      if get_inverse_kin_has_solution(pose.crt, qnear=pose.q):
          pose.jnt = get_inverse_kin(pose.crt, qnear=pose.q)
      else:
          popup("no solution found for the transition pose", blocking= True)
      end

      return pose
  end

  def get_transition_pose_2(ref, radius, axis_config, closest=False):
      # get the correspondig pose from the list of poses

      local jnt_current = get_actual_joint_positions()
      local yaw_current = get_yaw_too_base(ref)

      #pose.crt = get_tool_free_pose(pose_ref=ref, dir=[0, 0, DISTANCE_TO_CLEARANCE], move_in_base_frame=True)

      if (axis_config == 1):
          pose.q = JNT_STANDARD_C1
      elif (axis_config == 2):
          pose.q = JNT_STANDARD_C2
      end

      if closest:
          pose.q[0] = jnt_current[0]
      end

      # get coordinates of the circle with the same angle as the given pose to the
      if ref == p[0,0,0,0,0,0]:
          pose.crt = PSE_WA_1
      else:
          pose.crt =
          p[radius * cos(yaw_current-pi/2),
          radius * sin(yaw_current-pi/2),
          DISTANCE_TO_CLEARANCE,
          0,
          0,
          yaw_current + get_locked_yaw()]
      end

      if get_inverse_kin_has_solution(pose.crt, qnear=pose.q):
          pose.jnt = get_inverse_kin(pose.crt, qnear=pose.q)
          #return pose
      else:
          popup("no solution found for the transition pose", blocking= True)
      end

      return pose
  end

  def get_rounded_mm(value):
      if (value < 0):
          return ceil(value*1000)
      elif (value >= 0):
          return floor(value*1000)
      end
  end

  def get_yaw_too_base(pose):
      # get the yaw relative to the base frame
      local pose_x_mm = 0
      local pose_y_mm = 0
      local yaw = 0

      pose_x_mm = get_rounded_mm(pose[0])
      pose_y_mm = get_rounded_mm(pose[1])

      if (pose_x_mm == 0 and pose_y_mm < 0):
          yaw = 0
      elif (pose_x_mm == 0 and pose_y_mm > 0):
          yaw = pi
      elif (pose_x_mm < 0 and pose_y_mm == 0):
          yaw = -pi/2
      elif (pose_x_mm > 0 and pose_y_mm == 0):
          yaw = pi/2
      else:
          yaw = atan2(pose[0], pose[1])
          if (-pi < yaw) and (yaw < 0):
              yaw = - yaw - pi
          elif (0 < yaw) and (yaw < pi):
              yaw = - yaw + pi
          else:
              yaw = pi
          end
      end
      return yaw
  end

  def get_helper_pose():
      # get the helper pose, as described

      local m_line = 0                    # slope of the line between base and circle point
      local n = 0                         # shift on the ordinate axis
      local m_normal = 0                  # slope of the normal of the line between base and circle point
      local x_p1 = 0                      # x coordinate of first circle point
      local x_p2 = 0                      # x coordinate of second circle point
      local y_p1 = 0                      # y coordinate of first circle point
      local y_p2 = 0                      # y coordinate of second circle point
      local jnt_help_1 = [0,0,0,0,0,0]
      local jnt_help_2 = [0,0,0,0,0,0]

      if (pose_start.crt != pose_target.crt):
          if (pose_start.crt[0] == pose_target.crt[0]):
              m_normal = 0
          elif (pose_start.crt[0] != pose_target.crt[0]):
              m_line = (pose_target.crt[1]-pose_start.crt[1])/(pose_target.crt[0]-pose_start.crt[0])    # calculation of the slope between start and target
              n = pose_start.crt[1] - m_line * pose_start.crt[0]
          end
          if (-0.00001 > m_line or m_line > 0.00001):
              m_normal = -1/m_line
          end

          # using p-q-formula for getting the crossing points
          x_p1 = sqrt(pow(RADIUS_HELPER_POSES, 2)/(pow(m_normal, 2)+1)) * -1
          x_p2 = sqrt(pow(RADIUS_HELPER_POSES, 2)/(pow(m_normal, 2)+1))
          y_p1 = m_normal * x_p1
          y_p2 = m_normal * x_p2
          pose.q = pose_start.jnt

          if (point_dist(pose_start.crt, p[x_p1, y_p1,0,0,0,0]) < point_dist(pose_start.crt, p[x_p2, y_p2,0,0,0,0])):
              if reverse_rotation:
                  pose_help.crt[0] = x_p2
                  pose_help.crt[1] = y_p2
                  pose.q = pose_target.jnt
              else:
                  pose_help.crt[0] = x_p1
                  pose_help.crt[1] = y_p1
                  pose.q = pose_start.jnt
              end
          elif (point_dist(pose_start.crt, p[x_p1, y_p1,0,0,0,0]) > point_dist(pose_start.crt, p[x_p2, y_p2,0,0,0,0])):
              if reverse_rotation:
                  pose_help.crt[0] = x_p1
                  pose_help.crt[1] = y_p1
                  pose.q = pose_target.jnt
              else:
                  pose_help.crt[0] = x_p2
                  pose_help.crt[1] = y_p2
                  pose.q = pose_start.jnt
              end
          elif (point_dist(pose_start.crt, p[x_p1, y_p1,0,0,0,0]) == point_dist(pose_start.crt, p[x_p2, y_p2,0,0,0,0])):
              jnt_help_1 = get_inverse_kin(p[x_p1, y_p1,pose_start.crt[2],pose_start.crt[3],pose_start.crt[4],pose_start.crt[5]], qnear=pose.q)
              jnt_help_2 = get_inverse_kin(p[x_p2, y_p2,pose_start.crt[2],pose_start.crt[3],pose_start.crt[4],pose_start.crt[5]], qnear=pose.q)
              if (pose_start.jnt[0]<jnt_help_1[0] and jnt_help_1[0]<pose_target.jnt[0]) or (pose_start.jnt[0]>jnt_help_1[0] and jnt_help_1[0]>pose_target.jnt[0]):
                  pose_help.crt[0] = x_p1
                  pose_help.crt[1] = y_p1
              elif (pose_start.jnt[0]<jnt_help_2[0] and jnt_help_2[0]<pose_target.jnt[0]) or (pose_start.jnt[0]>jnt_help_2[0] and jnt_help_2[0]>pose_target.jnt[0]):
                  pose_help.crt[0] = x_p2
                  pose_help.crt[1] = y_p2
              end
              pose.q = pose_start.jnt
          end

          pose_help.crt[2] = 0.5 * (pose_start.crt[2] + pose_target.crt[2])

          if ((pose_start.crt[1] < 0 and pose_target.crt[1] > 0) or (pose_start.crt[1] > 0 and pose_target.crt[1] < 0)):
              if get_inverse_kin_has_solution(pose.crt, qnear=pose.q):
                  pose.jnt = get_inverse_kin(pose.crt, qnear=pose.q)
              else:
                  popup("no solution found for the helper pose", blocking= True)
              end
          end
      end
      return pose
  end

  def adjust_transition_poses(pose_identifier):
      # adjust the orientation of the transition poses by determining the the current orientation

      local pose_current = get_actual_tcp_pose()
      local jnt_current = get_actual_joint_positions()
      local rpy_current = rotvec2rpy([pose_current[3],pose_current[4],pose_current[5]])
      local rotvec_new = [0,0,0]

      if (pose_identifier == "start"):
          pose.q = pose_start.jnt
          pose.crt = get_forward_kin(pose_start.jnt)
      elif (pose_identifier == "helper"):
          pose.q = pose_help.jnt
          pose.crt = get_forward_kin(pose_help.jnt)
      elif (pose_identifier == "target"):
          pose.q = pose_target.jnt
          pose.crt = get_forward_kin(pose_target.jnt)
      end

      rotvec_new = rpy2rotvec([rpy_current[0], rpy_current[1], get_yaw_too_base(pose.crt) + yaw_locked])
      pose.crt = p[pose.crt[0], pose.crt[1], pose.crt[2], rotvec_new[0], rotvec_new[1], rotvec_new[2]]

      pose.q[3] = jnt_current[3]
      pose.q[4] = jnt_current[4]
      pose.q[5] = jnt_current[5]
      if get_inverse_kin_has_solution(pose.crt, qnear=pose.q) and is_within_safety_limits(pose.crt):
          pose.jnt = get_inverse_kin(pose.crt, qnear=pose.q)
      else:
          popup(str_cat("no solution for ", pose_identifier), error=True, blocking=True)
      end
      return pose.jnt
  end

  def get_locked_yaw():
      local pose_current = get_actual_tcp_pose()
      local rpy_current = rotvec2rpy([pose_current[3],pose_current[4],pose_current[5]])
      local rotvec_new = rpy2rotvec([rpy_current[0], rpy_current[1], get_yaw_too_base(pose_current)])
      local pose_reference = p[pose_current[0], pose_current[1], pose_current[2], rotvec_new[0], rotvec_new[1], rotvec_new[2]]
      local pose_to_reference = pose_trans(pose_inv(pose_reference), get_actual_tcp_pose())
      yaw_locked = pose_to_reference[5]

      return yaw_locked
  end

  def do_transition(reference_pose=p[0,0,0,0,0,0], mode=2, keep_xyz=[False, False, False], keep_rxry=False, a=1.4, v=1.05, r=0.100):
      # the robot will evaluate the current and target workarea
      # after that, the robot will move between the workareas automatically.
      # parameters:
      # reference_pose:   a pose/frame were the robot should work next. If nothing is given, base frame will be used as target
      # keep_rxry:        if true, the robot will keep the orientation of the tool during the movement

      ################# checking #################
      axis_config_current = check_current_axis_config()           # 0: unknown, 1: config 1, 2: config 2
      workarea_current = check_workarea(get_actual_tcp_pose())    # between 0 and the amount of defined workareas
      workarea_new = check_workarea(reference_pose)               # between 0 and the amount of defined workareas
      if(workarea_current==workarea_new):
           return 0
      end
      if (workarea_current != 0 and workarea_new != 0):
          ################# get axisvalues #################
          # pose_start = get_transition_pose(workarea_current, axis_config_current, closest=not reverse_rotation, keep_xyz=keep_xyz)
          pose_start = get_transition_pose_2(get_actual_tcp_pose(), RADIUS_TRANSITION_POSES, axis_config_current, closest=not reverse_rotation)
          if (workarea_current == 3 and workarea_new == 4) or (workarea_current == 4 and workarea_new == 3):
              # pose_target = get_transition_pose(workarea_new, axis_config_current, closest=True)
              pose_target = get_transition_pose_2(reference_pose, RADIUS_TRANSITION_POSES, axis_config_current, closest=True)
              reverse_rotation = True
          else:
              pose_target = get_transition_pose_2(reference_pose, RADIUS_TRANSITION_POSES, axis_config_current, closest=(workarea_current == workarea_new))
              if reverse_rotation:
                  reverse_rotation = False
              end
          end
          # pose_help = get_helper_pose()
          global A_Start = pose_start.crt
          global A_Help = pose_help.crt
          global A_End = pose_target.crt


          ################# adjustments #################
          if (keep_rxry):
              get_locked_yaw()
              if (pose_start.jnt == pose_target.jnt):
                  pose_target.jnt = adjust_transition_poses("target")
                  pose_start.jnt = pose_target.jnt
              else:
                  pose_start.jnt = adjust_transition_poses("start")
                  pose_target.jnt = adjust_transition_poses("target")
              end
              if (pose_help.jnt != [0,0,0,0,0,0]):
                  pose_help.jnt = adjust_transition_poses("helper")
              end
          end

          global A_Start = pose_start.crt
          global A_Help = pose_help.crt
          global A_End = pose_target.crt

          ################# movements #################

          if point_dist(pose_start.crt, pose_target.crt) > 0.100:
              movej(pose_start.jnt, a=a, v=v, r=r)
          end
          # if (pose_help.jnt != [0,0,0,0,0,0]):
          #     movej(pose_help.jnt, a=a, v=v, r=r)
          # end
          movej(pose_target.jnt, a=a, v=v)
      else:
          # define error
      end

      ################# checking #################
      axis_config_current = check_current_axis_config()           # 0: unknown, 1: config 1, 2: config 2
      workarea_current = check_workarea(get_actual_tcp_pose())    # between 0 and the amount of defined workareas
  end
  $ 5 "Script: SCRIPT Utility V5.1.script"
  #*****************************************************
  # customer          :   tbd
  # project name      :   tbd
  #****************************************************
  # controller        :
  # software          :
  #****************************************************
  # author            :   P. Koehnke (+49 1628859904; p.koehnke@unitedrobotics.group)
  # Copyright (c)     :   United Robotics Group Health and Food GmbH
  #                       An der Riede 2
  #                       28816 Stuhr
  #                       Germany
  #****************************************************
  # description       :   utility programs for the application
  # version:      	:   3.1
  # created           :   30.01.2023
  # updated           :
  #****************************************************
  # modifications     :   get_tool_free_pose_2(), get_index_from_list()
  #
  # date              :   05.01.2024
  # name              :   PK
  # reason            :
  #****************************************************

  def found_in_matrix(data, req_id, req_idx):
      local id = -1
      local dimensions = size(data)
      local loop_dataset = 0

      while (id != req_id and loop_dataset < dimensions[0]):
          id = data[loop_dataset, 0]
          if (id == req_id):
              return data[loop_dataset, req_idx]
          else:
              loop_dataset = loop_dataset + 1
          end
      end
  end

  def found_in_list(value, list):
      local idx = 0

      while (idx < length(list)):
          if (value == list[idx]):
              return True
          end
          idx = idx + 1
      end
      return False
  end

  def get_index_from_list(list, value=-1):
      local idx = 0

      while (idx < length(list)):
          if (value == -1):
              if (list[idx] != 0):
                  return idx
              end
          else:
              if (list[idx] == value):
                  return idx
              end
          end
          idx = idx + 1
      end
      return -1
  end

  def pose_RPY2RotVec(pose):
      local rotvec = rpy2rotvec([d2r(pose[3]),d2r(pose[4]),d2r(pose[5])])
      return p[pose[0],pose[1],pose[2],rotvec[0],rotvec[1],rotvec[2]]
  end

  def pose_RotVec2RPY(pose):
      local rpy = rotvec2rpy([pose[3],pose[4],pose[5]])
      return p[pose[0],pose[1],pose[2],r2d(rpy[0]),r2d(rpy[1]),r2d(rpy[2])]
  end

  def swivel(frame_ref, angles=[0,0,0], pose=p[0,0,0,0,0,0]):

      local rpy_ref = [0,0,0]
      local rpy_new = [0,0,0]
      local rotvec_new = [0,0,0]
      local pose_from = p[0,0,0,0,0,0]
      local pose_to = p[0,0,0,0,0,0]
      local i = 0

      if (pose == p[0,0,0,0,0,0]):
          pose_to = pose_trans(pose_inv(frame_ref), get_actual_tcp_pose())
      else:
          pose_to = pose
      end

      rpy_ref = rotvec2rpy(frame_ref[3], frame_ref[4], frame_ref[5])

      while (i < 3):
          rpy_new[i] = rpy_ref[i] + d2r(angles[i])
          i = i + 1
      end

      rotvec_new = rpy2rotvec(rpy_new)
      pose_from = p[0,0,0,rotvec_new[0],rotvec_new[1],rotvec_new[2]]
      pose_to = p[pose_to[0], pose_to[1], pose_to[2], rotvec_new[0], rotvec_new[1], rotvec_new[2]]

      return pose_trans(pose_from, pose_to)
  end

  def get_random_pose(pose_ref, mode="", range_max=[0,0,0]):
      # modi: "cubic", "rotation"
      # getting a random pose in the x/y-plane. range can be set for each
      # translation and rotation.
      local rpy_random = [0,0,0]
      local rotvec_random = [0,0,0]
      local pose_random = pose_ref
      local i = 0

      if (mode == "cubic"):
          # cubic mode: random pose takes only x, y and z
          i = 0
          while(i<3):
              pose_random[i] = pose_ref[i] + range_max[i] * (random() - 0.5)
              i = i + 1
          end
          return pose_random

      elif (mode == "rotation"):
          i = 0
          while(i<3):
              rpy_random[i] = d2r(range_max[i]) * (random() - 0.5)
              i = i + 1
          end
          rotvec_random = rpy2rotvec(rpy_random)
          pose_random = pose_trans(p[0,0,0,rotvec_random[0],rotvec_random[1],rotvec_random[2]], pose_ref)
          return pose_random

      else:
          # unknown mode, return pose_ref
          return pose_ref
      end
  end

  def get_pattern_pos_rectangle(counter, direction, patternsize, patterninc=[0,0], patternwidth=[0,0]):
      # defines the position inside a rectangular pattern
      # patternsize describes, how many objects are in x-direction and how many in y-direction [x, y]
      # patternwidth will give the total length of each direction [x, y]
      local X_Fac = 0
      local Y_Fac = 0
      local max = patternsize[0]*patternsize[1]

      if (1>counter or counter>max):
          counter = 1
      end

      if (direction == "Y" or direction == "y"):
          X_Fac = floor((counter - 1) / patternsize[1])
          Y_Fac = (counter - 1) % patternsize[1]
      elif (direction == "X" or direction == "x"):
          X_Fac = (counter - 1) % patternsize[0]
          Y_Fac = floor((counter - 1) / patternsize[0])
      end

      if patternwidth != [0,0]:
          patterninc = [patternwidth[0]/(patternsize[0]-1), patternwidth[1]/(patternsize[1]-1)]
      end

      return p[X_Fac*patterninc[0], Y_Fac*patterninc[1],0,0,0,0]
  end

  def get_pattern_pos_circle(counter, radius, angle, direction, pattern, patternsize=[0,0]):
      # get the patternpos for a circular pattern through a counter
      # need the radius and the angle in radiants
      local X_Fac = 0
      local Y_Fac = 0
      local rad_bow = 0
      local radius_cal = 0
      local ref = p[0,0,0,0,0,0]

      if (direction == "Y" or direction == "y"):
          X_Fac = floor((counter - 1) / pattern[1])
          Y_Fac = (counter - 1) % pattern[1]
      elif (direction == "X" or direction == "x"):
          X_Fac = (counter - 1) % pattern[0]
          Y_Fac = floor((counter - 1) / pattern[0])
      end

      # the opening angle will be calculated in x-direction
      # works only between -90 and 90 degree
      rad_bow = -angle/(pattern[0]-1) * X_Fac + angle/2

      if (counter%2 == 0):
          radius_cal = radius - patternsize[1]/(pattern[1])
      else:
          radius_cal = radius + patternsize[1]/(pattern[1])
      end
      ref = p[0, radius_cal, 0, 0, 0, 0]

      return p[ref[0]*cos(rad_bow)-ref[1]*sin(rad_bow), (ref[0]*sin(rad_bow)+ref[1]*cos(rad_bow))-radius,0,0,0,0]
  end

  def get_pattern_counter(pose, direction, pattern, patterninc=[0,0], patternsize=[0,0]):
      # returns the counter for a pattern from a given cartesian pose
      local patternpose = p[pose[0],pose[1],0,0,0,0]
      local floatFacX = 0.0
      local floatFacY = 0.0
      local remainder = 0.0
      local FacX = 0
      local FacY = 0

      # since the pattern spreads from the origin in positive axis-directions, all negative values
      # (which could appear due to a position near an axis) will set to zero
      if (pose[0]<0):
          patternpose = p[0,pose[1],0,0,0,0]
      end
      if (pose[1]<0):
          patternpose = p[pose[0],0,0,0,0,0]
      end
      # calculate the factor for each axis
      floatFacX = patternpose[0]/(patternsize[0]*(pattern[0]-1))
      floatFacY = patternpose[1]/(patternsize[1]*(pattern[1]-1))
      # determine the remainder after the comma/point
      if (floatFacX>1):
          remainder = floatFacX%floor(floatFacX)
      else:
          remainder = floatFacX
      end
      if (remainder<0.5):
          FacX = floatFacX-remainder
      else:
          FacX = floatFacX+(1-remainder)
      end

      if (floatFacY>1):
          remainder = floatFacY%floor(floatFacY)
      else:
          remainder = floatFacY
      end
      if (remainder<0.5):
          FacY = floatFacY-remainder
      else:
          FacY = floatFacY+(1-remainder)
      end
      # calculation of the counter in the desired axis-direction
      if (direction=="x" or direction=="X"):
          return FacX*pattern[1] + FacY + 1
      elif (direction=="y" or direction=="Y"):
          return FacY*pattern[0] + FacX + 1
      end
  end

  def get_plc_reg(mod_sig_name):
  	return integer_to_binary_list(modbus_get_signal_status(mod_sig_name))
  end

  def set_plc_reg(mod_sig_name, mod_sig_list):
  	modbus_set_output_register(mod_sig_name,binary_list_to_integer(mod_sig_list),False)
  end

  def check_decapping(offset=0, timeout=5):
      # checken, ob der Deckel schon ab ist
      local start = get_actual_tcp_pose()
      local current_offset = 0
      local timecounter = 0
      while (current_offset < offset):
          current_offset = pose_dist(start, get_actual_tcp_pose())
          timecounter = timecounter + 1
          if (timecounter*0.5 == timeout):
              break
          end
          sleep(0.5)
      end
      stopl(0.5)
  end

  def check_capping(torque=0):
      # checken, wann der Deckel verschraubt ist
      force_mode(get_actual_tcp_pose(), [0,0,1,0,0,0], [0,0,-2.0,0,0,0], 2, [0,0,0.100,0,0,0])
  end

  def is_reachable(frame, poses, offsets=[0,0,0]):
      local idx = 0
      local pose = p[0,0,0,0,0,0]

      while (idx < length(poses)):
          pose = poses[idx]
          pose[0] = pose[0] + offsets[0]
          pose[1] = pose[1] + offsets[1]
          pose[2] = pose[2] + offsets[2]

          if pose != p[0,0,0,0,0,0]:
              if (not get_inverse_kin_has_solution(pose_trans(frame, pose))):
                  textmsg(str_cat(str_cat("Pose ", to_str(idx + 1)), " is not reachable"))
                  return False
              end
          end
          idx = idx + 1
      end
      return True
  end

  def is_within_limits(frame, poses, offsets=[0,0,0]):
      local idx = 0
      local pose = p[0,0,0,0,0,0]

      while (idx < length(poses)):
          pose = poses[idx]
          pose[0] = pose[0] + offsets[0]
          pose[1] = pose[1] + offsets[1]
          pose[2] = pose[2] + offsets[2]

          if is_reachable(frame=frame, poses=poses, offsets=offsets):
              if (not is_within_safety_limits(get_inverse_kin(pose_trans(frame, pose), get_actual_joint_positions()))):
                  textmsg(str_cat(str_cat("Pose ", to_str(idx + 1)), "is out of joint limits"))
                  return False
              else:
                  idx = idx + 1
              end
          else:
              return False
          end
      end
      return True
  end

  def action_manipulator_decapping():
    zero_ftsensor()
    local DCP_Start = get_actual_tcp_pose ()
    global DCP_Actual = get_actual_tcp_pose ()
    local DCP_Height = 0.021
    global ForceCounter = 0
    sleep(0.02)
    zero_ftsensor()
    force_mode(p[0.0, 0.0, 0.0, 0.0, 0.0, 0.0], [0, 0, 1, 0, 0, 0], [0.0, 0.0, 17.0, 0.0, 0.0, 10.0], 2, [0.1, 0.1, 0.02, 0.3490658503988659, 0.3490658503988659, 0.3490658503988659])
    thread Thread_while_684():
      while (True):
        global DCP_Actual = get_actual_tcp_pose ()
        sleep(0.2)
        global ForceCounter = ForceCounter + 1
        if (ForceCounter > 30):
          zero_ftsensor()
          global ForceCounter = 0
        end
      end
    end
    if (DCP_Actual[2] <= DCP_Start[2] + DCP_Height):
      global thread_handler_decapping = run Thread_while_684()
      while (DCP_Actual[2] <= DCP_Start[2] + DCP_Height):
        sync()
      end
      kill thread_handler_decapping
    end
    end_force_mode()
    stopl(5.0)
  end
  $ 6 "PRC_Target≔0"
  global PRC_Target=0
  $ 7 "PRC_Target≔1"
  global PRC_Target=1
  $ 8 "Action≔1"
  global Action=1
  $ 9 "Action≔2"
  global Action=2
  $ 10 "Action≔7"
  global Action=7
  $ 11 "ITM_ID≔2"
  global ITM_ID=2
  $ 12 "JIG≔1"
  global JIG=1
  $ 13 "JIG_Slot≔2"
  global JIG_Slot=2
  $ 14 "Robot Program"
  $ 15 "PreSettings"
  $ 16 "init poses"
  $ 17 "PSE_A≔p[0,0,0,0,0,0]"
  global PSE_A=p[0,0,0,0,0,0]
  $ 18 "PSE_A_H≔p[0,0,0,0,0,0]"
  global PSE_A_H=p[0,0,0,0,0,0]
  $ 19 "PSE_T≔p[0,0,0,0,0,0]"
  global PSE_T=p[0,0,0,0,0,0]
  $ 20 "PSE_T_H≔p[0,0,0,0,0,0]"
  global PSE_T_H=p[0,0,0,0,0,0]
  $ 21 "PSE_G≔p[0,0,0,0,0,0]"
  global PSE_G=p[0,0,0,0,0,0]
  $ 22 "PSE_G_H≔p[0,0,0,0,0,0]"
  global PSE_G_H=p[0,0,0,0,0,0]
  $ 23 "PSE_R≔p[0,0,0,0,0,0]"
  global PSE_R=p[0,0,0,0,0,0]
  $ 24 "PSE_R_H≔p[0,0,0,0,0,0]"
  global PSE_R_H=p[0,0,0,0,0,0]
  $ 25 "JNT_A≔[0,0,0,0,0,0]"
  global JNT_A=[0,0,0,0,0,0]
  $ 26 "JNT_S≔[0,0,0,0,0,0]"
  global JNT_S=[0,0,0,0,0,0]
  $ 27 "PROCESS_Info≔'work at target, Table'"
  global PROCESS_Info="work at target, Table"
  $ 28 "PRM_TubHghtDiff≔-0.024"
  global PRM_TubHghtDiff=-0.024
  $ 29 "Gripping parameters"
  $ 30 "GRP_Open_Pos≔45"
  global GRP_Open_Pos=45
  $ 31 "GRP_Close_Pos≔100"
  global GRP_Close_Pos=100
  $ 32 "rq_set_force_norm(20)"
   rq_set_force_norm (20)
  $ 33 "rq_set_speed_norm(80)"
   rq_set_speed_norm (80)
  $ 34 "Switch ITM_ID"
  switch_1 = ITM_ID
  $ 35 "Case 1"
  if (1 == switch_1):
    $ 36 "uML"
    $ 37 "Switch JIG"
    switch_2 = JIG
    $ 38 "Case 2"
    if (2 == switch_2):
      $ 39 "biorad rack tubes"
      $ 40 "GRP_Open_Pos≔60"
      global GRP_Open_Pos=60
      $ 41 "FRM_Reference≔uLM_BradRckTubs"
      global FRM_Reference=uLM_BradRckTubs
      $ 42 "PSE_T≔pose_RPY2RotVec(p[0.02*(JIG_Slot%10),-0.0334*floor(JIG_Slot/10),0,0,0,-90])"
      global PSE_T=pose_RPY2RotVec(p[0.02*(JIG_Slot%10),-0.0334*floor(JIG_Slot/10),0,0,0,-90])
      $ 43 "PSE_T[2]=PSE_T[2]+PRM_TubHghtDiff"
      PSE_T[2]=PSE_T[2]+PRM_TubHghtDiff
      $ 44 "If (JIG_Slot%10)>1"
      if ((JIG_Slot%10)>1):
        $ 45 "PSE_T[0]=PSE_T[0]+0.0165"
        PSE_T[0]=PSE_T[0]+0.0165
        $ 46 "If (JIG_Slot%10)>4"
        if ((JIG_Slot%10)>4):
          $ 47 "PSE_T[0]=PSE_T[0]+0.0235"
          PSE_T[0]=PSE_T[0]+0.0235
          $ 48 "If (JIG_Slot%10)>6"
          if ((JIG_Slot%10)>6):
            $ 49 "PSE_T[0]=PSE_T[0]+0.0165"
            PSE_T[0]=PSE_T[0]+0.0165
          end
        end
      end
      $ 50 "PSE_R≔pose_add(PSE_T, p[0,0,0.2500,0,0,0])"
      global PSE_R= pose_add (PSE_T, p[0,0,0.2500,0,0,0])
      $ 51 "PSE_A≔pose_add(PSE_T, p[0,0,0.1,0,0,0])"
      global PSE_A= pose_add (PSE_T, p[0,0,0.1,0,0,0])
    elif (4 == switch_2):
      $ 52 "Case 4"
      $ 53 "centrifuge rack tubes"
      $ 54 "GRP_Open_Pos≔60"
      global GRP_Open_Pos=60
      $ 55 "FRM_Reference≔uLM_CentTubes"
      global FRM_Reference=uLM_CentTubes
      $ 56 "PSE_T≔pose_RPY2RotVec(p[0.0975*(JIG_Slot%4),0,0,0,0,0])"
      global PSE_T=pose_RPY2RotVec(p[0.0975*(JIG_Slot%4),0,0,0,0,0])
      $ 57 "PSE_T[2]=PSE_T[2]+PRM_TubHghtDiff"
      PSE_T[2]=PSE_T[2]+PRM_TubHghtDiff
      $ 58 "If JIG_Slot>3 and JIG_Slot≤7"
      if (JIG_Slot>3  and  JIG_Slot <= 7):
        $ 59 "PSE_T[1]=0.06"
        PSE_T[1]=0.06
        $ 60 "PSE_T[0]=PSE_T[0]+0.06"
        PSE_T[0]=PSE_T[0]+0.06
      else:
        $ 61 "ElseIf JIG_Slot>7 and JIG_Slot≤11"
        if (JIG_Slot>7  and  JIG_Slot <= 11):
          $ 62 "PSE_T[0]=PSE_T[0]+0.06"
          PSE_T[0]=PSE_T[0]+0.06
        else:
          $ 63 "ElseIf JIG_Slot>11 and JIG_Slot≤15"
          if (JIG_Slot>11  and  JIG_Slot <= 15):
            $ 64 "PSE_T[1]=0.06"
            PSE_T[1]=0.06
          end
        end
      end
      $ 65 "PSE_R≔pose_add(PSE_T, p[0,0,0.150,0,0,0])"
      global PSE_R= pose_add (PSE_T, p[0,0,0.150,0,0,0])
      $ 66 "PSE_A≔pose_add(PSE_T, p[0,0,0.15,0,0,0])"
      global PSE_A= pose_add (PSE_T, p[0,0,0.15,0,0,0])
    elif (5 == switch_2):
      $ 67 "Case 5"
      $ 68 "3finger gripper"
      $ 69 "define poses"
      $ 70 "'Place in 3finger'"
      # 'Place in 3finger'
      $ 71 "FRM_Reference = uML_3fingergrip"
      FRM_Reference = uML_3fingergrip
      $ 72 "PSE_T≔pose_RPY2RotVec(p[0,0,0.002,0,0,0])"
      global PSE_T=pose_RPY2RotVec(p[0,0,0.002,0,0,0])
      $ 73 "PSE_T[2]=PSE_T[2]+PRM_TubHghtDiff"
      PSE_T[2]=PSE_T[2]+PRM_TubHghtDiff
      $ 74 "If Action≟5"
      if (Action == 5):
        $ 75 "PSE_T≔pose_RPY2RotVec(p[0,0,0.018,0,0,0])"
        global PSE_T=pose_RPY2RotVec(p[0,0,0.018,0,0,0])
        $ 76 "PSE_T_H≔pose_trans(PSE_T, p[0,0,0.02,0,0,0])"
        global PSE_T_H= pose_trans (PSE_T, p[0,0,0.02,0,0,0])
      end
      $ 77 "If Action≟3"
      if (Action == 3):
        $ 78 "PSE_T[5]=PSE_T[5]+d2r(155)"
        PSE_T[5]=PSE_T[5]+d2r(155)
      end
      $ 79 "PSE_A≔pose_trans(PSE_T, p[0,0,0.1,0,0,0])"
      global PSE_A= pose_trans (PSE_T, p[0,0,0.1,0,0,0])
      $ 80 "PSE_R≔pose_add(PSE_T, p[0,0,0.060,0,0,0])"
      global PSE_R= pose_add (PSE_T, p[0,0,0.060,0,0,0])
    elif (6 == switch_2):
      $ 81 "Case 6"
      $ 82 "Caps bin"
      $ 83 "define poses"
      $ 84 "'Drop cap'"
      # 'Drop cap'
      $ 85 "FRM_Reference=uML_CapBin"
      FRM_Reference=uML_CapBin
      $ 86 "PSE_T≔pose_RPY2RotVec(p[0,0,0,0,0,0])"
      global PSE_T=pose_RPY2RotVec(p[0,0,0,0,0,0])
      $ 87 "PSE_T_H≔pose_trans(PSE_T, p[0,0,-0.006,0,0,0])"
      global PSE_T_H= pose_trans (PSE_T, p[0,0,-0.006,0,0,0])
      $ 88 "PSE_A≔pose_trans(PSE_T, p[0,0,0.1,0,0,0])"
      global PSE_A= pose_trans (PSE_T, p[0,0,0.1,0,0,0])
      $ 89 "PSE_R≔pose_add(PSE_T, p[0,0,0.100,0,0,0])"
      global PSE_R= pose_add (PSE_T, p[0,0,0.100,0,0,0])
    elif (7 == switch_2):
      $ 90 "Case 7"
      $ 91 "define poses Manual"
      $ 92 "GRP_Open_Pos≔60"
      global GRP_Open_Pos=60
      $ 93 "FRM_Reference≔uLM_Manual"
      global FRM_Reference=uLM_Manual
      $ 94 "If Action≟1"
      if (Action == 1):
        $ 96 "PSE_T≔pose_RPY2RotVec(p[0.0248*(JIG_Slot%8),0.0258*(floor(JIG_Slot/8)),0,0,0,0])"
        global PSE_T=pose_RPY2RotVec(p[0.0248*(JIG_Slot%8),0.0258*(floor(JIG_Slot/8)),0,0,0,0])
        $ 97 "PSE_R≔pose_add(PSE_T, p[0,0,0.2500,0,0,0])"
        global PSE_R= pose_add (PSE_T, p[0,0,0.2500,0,0,0])
      else:
        $ 98 "ElseIf Action≟2"
        if (Action == 2):
          $ 100 "PSE_T≔pose_RPY2RotVec(p[0.0248*(JIG_Slot%8),0.0258*(floor(JIG_Slot/8)),0,0,0,0])"
          global PSE_T=pose_RPY2RotVec(p[0.0248*(JIG_Slot%8),0.0258*(floor(JIG_Slot/8)),0,0,0,0])
          $ 101 "PSE_R≔pose_add(PSE_T, p[0,0,0.100,0,0,0])"
          global PSE_R= pose_add (PSE_T, p[0,0,0.100,0,0,0])
        end
      end
      $ 102 "PSE_T[2]=PSE_T[2]+PRM_TubHghtDiff"
      PSE_T[2]=PSE_T[2]+PRM_TubHghtDiff
      $ 103 "PSE_A≔pose_add(PSE_T, p[0,0,0.1,0,0,0])"
      global PSE_A= pose_add (PSE_T, p[0,0,0.1,0,0,0])
    end
  elif (2 == switch_1):
    $ 104 "Case 2"
    $ 105 "Biorad"
    $ 106 "'CHANGE THE REFERENCE TO THE FRAME TO MOVE IN'"
    # 'CHANGE THE REFERENCE TO THE FRAME TO MOVE IN'
    $ 107 "Gripping parameters"
    $ 108 "GRP_Open_Pos≔45"
    global GRP_Open_Pos=45
    $ 109 "GRP_Close_Pos≔100"
    global GRP_Close_Pos=100
    $ 110 "rq_set_force_norm(80)"
     rq_set_force_norm (80)
    $ 111 "rq_set_speed_norm(100)"
     rq_set_speed_norm (100)
    $ 112 "If PRC_Target≟0"
    if (PRC_Target == 0):
      $ 113 "FRM_Reference = uML_BradRacks"
      FRM_Reference = uML_BradRacks
      $ 114 "PSE_T≔pose_RPY2RotVec(p[0.0347*JIG_Slot,0,0,0,0,180])"
      global PSE_T=pose_RPY2RotVec(p[0.0347*JIG_Slot,0,0,0,0,180])
      $ 115 "PSE_A≔pose_add(PSE_T, p[0,0,0.18,0,0,0])"
      global PSE_A= pose_add (PSE_T, p[0,0,0.18,0,0,0])
      $ 116 "PSE_R≔pose_add(PSE_T, p[0,0,0.18,0,0,0])"
      global PSE_R= pose_add (PSE_T, p[0,0,0.18,0,0,0])
    else:
      $ 117 "Else" "noBreak"
      $ 118 "FRM_Reference = FRM_BioradMachn"
      FRM_Reference = FRM_BioradMachn
      $ 119 "If Action≟7"
      if (Action == 7):
        $ 120 "PSE_T≔pose_RPY2RotVec(p[0.125-0.056*JIG_Slot,0.084,0.028,-72,0,0])"
        global PSE_T=pose_RPY2RotVec(p[0.125-0.056*JIG_Slot,0.084,0.028,-72,0,0])
        $ 121 "PSE_T_H≔pose_RPY2RotVec(p[0.126-0.056*JIG_Slot,0.084,0.254,-72,0,0])"
        global PSE_T_H=pose_RPY2RotVec(p[0.126-0.056*JIG_Slot,0.084,0.254,-72,0,0])
        $ 122 "PSE_A≔pose_add(PSE_T_H, p[0,0.1,0,0,0,0])"
        global PSE_A= pose_add (PSE_T_H, p[0,0.1,0,0,0,0])
        $ 123 "PSE_R≔pose_add(PSE_T_H, p[0,0.1,0.1,0,0,0])"
        global PSE_R= pose_add (PSE_T_H, p[0,0.1,0.1,0,0,0])
      else:
        $ 124 "ElseIf Action≟2"
        if (Action == 2):
          $ 125 "PSE_T≔pose_RPY2RotVec(p[0.126-0.056*JIG_Slot,0.07,0.08,-90,0,0])"
          global PSE_T=pose_RPY2RotVec(p[0.126-0.056*JIG_Slot,0.07,0.08,-90,0,0])
          $ 126 "PSE_T_H≔pose_RPY2RotVec(p[0.126-0.056*JIG_Slot,0.072,0.238,-90,0,0])"
          global PSE_T_H=pose_RPY2RotVec(p[0.126-0.056*JIG_Slot,0.072,0.238,-90,0,0])
          $ 127 "PSE_A≔pose_add(PSE_T_H, p[0,0.1,0,0,0,0])"
          global PSE_A= pose_add (PSE_T_H, p[0,0.1,0,0,0,0])
          $ 128 "PSE_R≔pose_add(PSE_T_H, p[0,0.1,0,0,0,0])"
          global PSE_R= pose_add (PSE_T_H, p[0,0.1,0,0,0,0])
        end
      end
    end
  elif (4 == switch_1):
    $ 132 "Case 4"
    $ 133 "Centrifuge"
    $ 134 "'CHANGE THE REFERENCE TO THE FRAME TO MOVE IN'"
    # 'CHANGE THE REFERENCE TO THE FRAME TO MOVE IN'
    $ 135 "Gripping parameters"
    $ 136 "GRP_Open_Pos≔45"
    global GRP_Open_Pos=45
    $ 137 "GRP_Close_Pos≔100"
    global GRP_Close_Pos=100
    $ 138 "rq_set_force_norm(80)"
     rq_set_force_norm (80)
    $ 139 "rq_set_speed_norm(100)"
     rq_set_speed_norm (100)
    $ 140 "If PRC_Target≟0"
    if (PRC_Target == 0):
      $ 141 "FRM_Reference = uLM_CentRacks"
      FRM_Reference = uLM_CentRacks
    else:
      $ 142 "Else" "noBreak"
      $ 143 "FRM_Reference = FRM_Centrifuge"
      FRM_Reference = FRM_Centrifuge
    end
    $ 144 "PSE_T≔pose_RPY2RotVec(p[0,0,0,0,0,0])"
    global PSE_T=pose_RPY2RotVec(p[0,0,0,0,0,0])
    $ 145 "PSE_A≔pose_add(PSE_T, p[0,0,0.1,0,0,0])"
    global PSE_A= pose_add (PSE_T, p[0,0,0.1,0,0,0])
    $ 146 "PSE_R≔pose_add(PSE_T, p[0,0,0.1,0,0,0])"
    global PSE_R= pose_add (PSE_T, p[0,0,0.1,0,0,0])
  end
  $ 147 "Additional check"
  $ 148 "If  not is_reachable(FRM_Reference,[PSE_A,PSE_A_H,PSE_T,PSE_T_H,PSE_R,PSE_R_H])"
  if (  not  is_reachable(FRM_Reference,[PSE_A,PSE_A_H,PSE_T,PSE_T_H,PSE_R,PSE_R_H])):
    $ 149 "set_error(1002)"
    set_error(1002)
    $ 150 "Action≔0"
    global Action=0
  end
  $ 151 "Switch Action"
  switch_1 = Action
  $ 152 "Case 1"
  if (1 == switch_1):
    $ 153 "Pick"
    $ 154 "Action_Info≔'Pick Rack/Probe'"
    global Action_Info="Pick Rack/Probe"
    $ 155 "do_transition(FRM_Reference, keep_rxry=OBJ_Picked)"
    do_transition(FRM_Reference, keep_rxry=OBJ_Picked)
    $ 156 "If  not OBJ_Picked"
    if (  not  OBJ_Picked):
      $ 157 "rq_move_and_wait_norm(GRP_Open_Pos)"
       rq_move_and_wait_norm (GRP_Open_Pos)
    end
    $ 158 "If JNT_A≠[0,0,0,0,0,0]"
    if (JNT_A != [0,0,0,0,0,0]):
      $ 159 "MoveJ"
      $ 160 "JNT_A" "breakAfter"
      movej(JNT_A, a=1.3962634015954636, v=1.7453292519943295, r=0.02)
    else:
      $ 161 "Else" "noBreak"
      $ 162 "MoveJ"
      $ 163 "PSE_A" "breakAfter"
      movej(pose_trans(FRM_Reference, PSE_A), a=1.3962634015954636, v=1.7453292519943295, r=0.02)
    end
    $ 164 "MoveL"
    $ 165 "PSE_T" "breakAfter"
    movel(pose_trans(FRM_Reference, PSE_T), a=0.08, v=0.12)
    $ 166 "rq_set_force_norm(50)"
     rq_set_force_norm (50)
    $ 167 "rq_move_and_wait_norm(GRP_Close_Pos)"
     rq_move_and_wait_norm (GRP_Close_Pos)
    $ 168 "OBJ_Picked≔rq_is_object_detected()"
    global OBJ_Picked= rq_is_object_detected ()
    $ 169 "If PSE_T_H≠PSE_Z"
    if (PSE_T_H != PSE_Z):
      $ 170 "PSE_T_H" "breakAfter"
      movel(pose_trans(FRM_Reference, PSE_T_H), a=0.5, v=0.4, r=0.01)
    end
    $ 171 "PSE_R" "breakAfter"
    movel(pose_trans(FRM_Reference, PSE_R), a=0.5, v=0.4)
  elif (2 == switch_1):
    $ 172 "Case 2"
    $ 173 "Place"
    $ 174 "Action_Info≔'place object'"
    global Action_Info="place object"
    $ 175 "do_transition(keep_rxry=OBJ_Picked)"
    do_transition(keep_rxry=OBJ_Picked)
    $ 176 "If JNT_A≠[0,0,0,0,0,0]"
    if (JNT_A != [0,0,0,0,0,0]):
      $ 177 "MoveJ"
      $ 178 "JNT_A" "breakAfter"
      movej(JNT_A, a=1.3962634015954636, v=1.7453292519943295, r=0.02)
    else:
      $ 179 "Else" "noBreak"
      $ 180 "MoveJ"
      $ 181 "PSE_A" "breakAfter"
      movej(pose_trans(FRM_Reference, PSE_A), a=1.3962634015954636, v=1.7453292519943295, r=0.02)
    end
    $ 182 "MoveL"
    $ 183 "If PSE_T_H≠PSE_Z"
    if (PSE_T_H != PSE_Z):
      $ 184 "PSE_T_H" "breakAfter"
      movel(pose_trans(FRM_Reference, PSE_T_H), a=0.04, v=0.07)
    end
    $ 185 "If JIG≟4 or ITM_ID≟2"
    if (JIG == 4  or  ITM_ID == 2):
      $ 186 "PSE_T" "breakAfter"
      movel(pose_trans(FRM_Reference, PSE_T), a=0.05, v=0.09)
    else:
      $ 187 "Else" "noBreak"
      $ 188 "PSE_T" "breakAfter"
      global move_thread_flag_188=0
      thread move_thread_188():
        enter_critical
        move_thread_flag_188 = 1
        movel(pose_trans(FRM_Reference, PSE_T), a=0.05, v=0.09)
        move_thread_flag_188 = 2
        exit_critical
      end
      move_thread_flag_188 = 0
      move_thread_han_188 = run move_thread_188()
      while (True):
        local targetTcpDirection=get_target_tcp_speed()
        local stepsToRetract=tool_contact(direction=targetTcpDirection)
        if (stepsToRetract > 0):
          kill move_thread_han_188
          stopl(0.5)
          local backTrackMovement=get_actual_joint_positions_history(stepsToRetract)
          local contactPose=get_forward_kin(backTrackMovement)
          local posDir=[targetTcpDirection[0],targetTcpDirection[1],targetTcpDirection[2]]
          local retractTo=contactPose
          if (norm(posDir) > 1e-6):
            local normalizedPosDir=normalize(posDir)
            local additionalRetraction=p[normalizedPosDir[0] * 0.0, normalizedPosDir[1] * 0.0, normalizedPosDir[2] * 0.0, 0, 0, 0]
            retractTo = pose_sub(contactPose, additionalRetraction)
          end
          movel(retractTo, a=0.5, v=0.1)
          $ 189 "Until (tool_contact_detection)"
          break
        end
        sleep(1.0E-10)
        if (move_thread_flag_188 > 1):
          join move_thread_han_188
          break
        end
        sync()
      end
      $ 190 "Force"
      sleep(0.02)
      zero_ftsensor()
      force_mode(FRM_Reference, [1, 1, 0, 0, 0, 0], [0.0, 0.0, 0.0, 0.0, 0.0, 0.0], 2, [0.05, 0.05, 0.1, 0.3490658503988659, 0.3490658503988659, 0.3490658503988659])
      $ 191 "PSE_T" "noBreak"
      movel(pose_trans(FRM_Reference, PSE_T), a=0.04, v=0.07)
      end_force_mode()
      stopl(5.0)
    end
    $ 192 "'ADD OPEN GRIPPER'"
    # 'ADD OPEN GRIPPER'
    $ 193 "rq_move_and_wait_norm(GRP_Open_Pos)"
     rq_move_and_wait_norm (GRP_Open_Pos)
    $ 194 "Wait: 0.2"
    sleep(0.2)
    $ 195 "PSE_R" "breakAfter"
    movel(pose_trans(FRM_Reference, PSE_R), a=0.5, v=0.4)
  elif (3 == switch_1):
    $ 197 "Case 3"
    $ 198 "Pick decapped probe from 3finger"
    $ 199 "Action_Info≔'Pick Rack/Probe'"
    global Action_Info="Pick Rack/Probe"
    $ 200 "MoveJ"
    $ 201 "PSE_A" "breakAfter"
    movej(pose_trans(FRM_Reference, PSE_A), a=1.3962634015954636, v=1.7453292519943295)
    $ 202 "rq_move_and_wait_norm(GRP_Open_Pos)"
     rq_move_and_wait_norm (GRP_Open_Pos)
    $ 203 "MoveL"
    $ 205 "PSE_T" "breakAfter"
    movel(pose_trans(FRM_Reference, PSE_T), a=0.15, v=0.075)
    $ 208 "'ADD OPEN GRIPPER'"
    # 'ADD OPEN GRIPPER'
    $ 209 "rq_set_force_norm(20)"
     rq_set_force_norm (20)
    $ 210 "rq_set_speed_norm(30)"
     rq_set_speed_norm (30)
    $ 211 "rq_move_and_wait_norm(GRP_Close_Pos)"
     rq_move_and_wait_norm (GRP_Close_Pos)
    $ 212 "Set Open3FG=On"
    set_standard_digital_out(4, True)
    $ 213 "Wait: 0.3"
    sleep(0.3)
    $ 214 "MoveL"
    $ 215 "PSE_R" "breakAfter"
    movel(pose_trans(FRM_Reference, PSE_R), a=1.2, v=0.25)
  elif (4 == switch_1):
    $ 216 "Case 4"
    $ 217 "Place probe in 3finger"
    $ 218 "Action_Info≔'place object'"
    global Action_Info="place object"
    $ 219 "MoveJ"
    $ 220 "PSE_A" "breakAfter"
    movej(pose_trans(FRM_Reference, PSE_A), a=1.3962634015954636, v=1.7453292519943295)
    $ 221 "Set Open3FG=On"
    set_standard_digital_out(4, True)
    $ 222 "MoveL"
    $ 223 "PSE_T" "breakAfter"
    global move_thread_flag_223=0
    thread move_thread_223():
      enter_critical
      move_thread_flag_223 = 1
      movel(pose_trans(FRM_Reference, PSE_T), a=0.15, v=0.075)
      move_thread_flag_223 = 2
      exit_critical
    end
    move_thread_flag_223 = 0
    move_thread_han_223 = run move_thread_223()
    while (True):
      local targetTcpDirection=get_target_tcp_speed()
      local stepsToRetract=tool_contact(direction=targetTcpDirection)
      if (stepsToRetract > 0):
        kill move_thread_han_223
        stopl(3.0)
        local backTrackMovement=get_actual_joint_positions_history(stepsToRetract)
        local contactPose=get_forward_kin(backTrackMovement)
        local posDir=[targetTcpDirection[0],targetTcpDirection[1],targetTcpDirection[2]]
        local retractTo=contactPose
        if (norm(posDir) > 1e-6):
          local normalizedPosDir=normalize(posDir)
          local additionalRetraction=p[normalizedPosDir[0] * 0.0, normalizedPosDir[1] * 0.0, normalizedPosDir[2] * 0.0, 0, 0, 0]
          retractTo = pose_sub(contactPose, additionalRetraction)
        end
        movel(retractTo, a=3.0, v=0.1)
        $ 224 "Until (tool_contact_detection)"
        break
      end
      sleep(1.0E-10)
      if (move_thread_flag_223 > 1):
        join move_thread_han_223
        break
      end
      sync()
    end
    $ 225 "Set Open3FG=Off"
    set_standard_digital_out(4, False)
    $ 226 "Wait: 0.5"
    sleep(0.5)
  elif (5 == switch_1):
    $ 231 "Case 5"
    $ 248 "Decapping"
    $ 249 "Action_Info≔'decapping'"
    global Action_Info="decapping"
    $ 250 "Set EN_3FG=On"
    set_standard_digital_out(5, True)
    $ 251 "Set DecapTurn=On"
    set_standard_digital_out(3, True)
    $ 252 "action_manipulator_decapping()"
    action_manipulator_decapping()
    $ 253 "Set EN_3FG=Off"
    set_standard_digital_out(5, False)
    $ 254 "Set DecapTurn=Off"
    set_standard_digital_out(3, False)
    $ 255 "MoveL"
    $ 256 "PSE_R" "breakAfter"
    movel(pose_trans(FRM_Reference, PSE_R), a=0.8, v=0.15)
  elif (6 == switch_1):
    $ 257 "Case 6"
    $ 276 "Drop"
    $ 277 "rq_set_speed_norm(100)"
     rq_set_speed_norm (100)
    $ 278 "MoveJ"
    $ 279 "PSE_A" "breakAfter"
    movej(pose_trans(FRM_Reference, PSE_A), a=1.3962634015954636, v=1.7453292519943295, r=0.02)
    $ 280 "MoveL"
    $ 281 "PSE_T" "breakAfter"
    movel(pose_trans(FRM_Reference, PSE_T), a=0.08, v=0.12)
    # begin: URCap Program Node
    #   Source: Robotiq_Grippers, 3.11.2.92906, Robotiq Inc.
    #   Type: Gripper
    $ 282 "Gripper Move14mm (1)"
    if not(gripper_connected[0]):
      popup("Gripper 1 must be connected to run this program.", "No connection", False, True, True)
    end
    if not(rq_is_gripper_activated("1")):
      popup("Gripper 1 is not activated. Go to Installation tab > Gripper to activate it and run the program again.", "Not activated", False, True, True)
    end
    rq_set_pos_spd_for(153, 255, 77, "1")
    rq_wait_pos_spe_for_request(153, 255, 77, "1")
    rq_go_to("1")
    rq_wait("1")
    # end: URCap Program Node
    $ 283 "PSE_T_H" "breakAfter"
    movel(pose_trans(FRM_Reference, PSE_T_H), a=0.08, v=0.12)
    $ 284 "rq_move_and_wait_norm(GRP_Open_Pos)"
     rq_move_and_wait_norm (GRP_Open_Pos)
    $ 285 "Wait: 0.2"
    sleep(0.2)
    $ 286 "PSE_R" "breakAfter"
    movel(pose_trans(FRM_Reference, PSE_R), a=0.5, v=0.4)
  elif (7 == switch_1):
    $ 287 "Case 7"
    $ 288 "Load"
    $ 289 "Action_Info≔'load object in the machine'"
    global Action_Info="load object in the machine"
    $ 291 "If JNT_A≠[0,0,0,0,0,0]"
    if (JNT_A != [0,0,0,0,0,0]):
      $ 292 "MoveJ"
      $ 293 "JNT_A" "breakAfter"
      movej(JNT_A, a=1.3962634015954636, v=1.7453292519943295, r=0.02)
    else:
      $ 294 "Else" "noBreak"
      $ 295 "MoveJ"
      $ 296 "PSE_A" "breakAfter"
      movej(pose_trans(FRM_Reference, PSE_A), a=1.3962634015954636, v=1.7453292519943295, r=0.02)
    end
    $ 297 "MoveL"
    $ 302 "PSE_T_H" "breakAfter"
    movel(pose_trans(FRM_Reference, PSE_T_H), a=0.04, v=0.07)
    $ 303 "rq_move_and_wait_norm(GRP_Close_Pos)"
     rq_move_and_wait_norm (GRP_Close_Pos)
    $ 304 "Wait: 0.2"
    sleep(0.2)
    $ 305 "PSE_T" "breakAfter"
    movel(pose_trans(FRM_Reference, PSE_T), a=0.04, v=0.07)
    # begin: URCap Program Node
    #   Source: Robotiq_Grippers, 3.11.2.92906, Robotiq Inc.
    #   Type: Gripper
    $ 306 "Gripper Move18mm (1)"
    if not(gripper_connected[0]):
      popup("Gripper 1 must be connected to run this program.", "No connection", False, True, True)
    end
    if not(rq_is_gripper_activated("1")):
      popup("Gripper 1 is not activated. Go to Installation tab > Gripper to activate it and run the program again.", "Not activated", False, True, True)
    end
    rq_set_pos_spd_for(127, 0, 173, "1")
    rq_wait_pos_spe_for_request(127, 0, 173, "1")
    rq_go_to("1")
    rq_wait("1")
    # end: URCap Program Node
    $ 307 "PSE_R" "breakAfter"
    movel(pose_trans(FRM_Reference, PSE_R), a=0.5, v=0.4)
  elif (16 == switch_1):
    $ 308 "Case 16"
    $ 309 "Scan the barcode"
    $ 310 "Action_Info≔'scan the barcode'"
    global Action_Info="scan the barcode"
    $ 311 "Barc_scan_succs≔ False "
    global Barc_scan_succs=  False
    $ 312 "First check"
    $ 313 "Set BarcodeTrigger=On"
    set_standard_digital_out(6, True)
    $ 314 "Wait: 0.1"
    sleep(0.1)
    $ 315 "Barc_scan_succs≔BarcodeSignal"
    global Barc_scan_succs=get_standard_digital_in(6)
    $ 316 "If Barc_scan_succs"
    if (Barc_scan_succs):
      $ 317 "Set EN_3FG=On"
      set_standard_digital_out(5, True)
      $ 318 "Set CapTurn=On"
      set_standard_digital_out(2, True)
      $ 319 "Loop Barc_scan_succs"
      thread Thread_while_319():
        while (True):
          $ 320 "Barc_scan_succs≔BarcodeSignal"
          global Barc_scan_succs=get_standard_digital_in(6)
          $ 321 "Wait: 0.05"
          sleep(0.05)
        end
      end
      if (Barc_scan_succs):
        global thread_handler_319=run Thread_while_319()
        while (Barc_scan_succs):
          sync()
        end
        kill thread_handler_319
      end
      $ 322 "Set EN_3FG=Off"
      set_standard_digital_out(5, False)
      $ 323 "Set CapTurn=Off"
      set_standard_digital_out(2, False)
      $ 324 "Set BarcodeTrigger=Off"
      set_standard_digital_out(6, False)
    else:
      $ 325 "Else" "noBreak"
      $ 326 "Timer_Barc_scan: Reset"
      Timer_Barc_scan = 0
      $ 327 "Timer_Barc_scan: Start"
      Timer_Barc_scan_is_counting = True
      $ 328 "Set DecapTurn=On"
      set_standard_digital_out(3, True)
      $ 329 "Set EN_3FG=On"
      set_standard_digital_out(5, True)
      $ 330 "Loop  not Barc_scan_succs and  not CMD_Stop and Timer_Barc_scan<60"
      thread Thread_while_330():
        while (True):
          $ 333 "Set BarcodeTrigger=On"
          set_standard_digital_out(6, True)
          $ 334 "Barc_scan_succs≔BarcodeSignal"
          global Barc_scan_succs=get_standard_digital_in(6)
          $ 335 "Wait: 0.05"
          sleep(0.05)
        end
      end
      if (  not  Barc_scan_succs  and    not  CMD_Stop  and  Timer_Barc_scan<60):
        global thread_handler_330=run Thread_while_330()
        while (  not  Barc_scan_succs  and    not  CMD_Stop  and  Timer_Barc_scan<60):
          sync()
        end
        kill thread_handler_330
      end
      $ 336 "Set EN_3FG=Off"
      set_standard_digital_out(5, False)
      $ 337 "Set DecapTurn=Off"
      set_standard_digital_out(3, False)
      $ 338 "Set BarcodeTrigger=Off"
      set_standard_digital_out(6, False)
      $ 339 "Timer_Barc_scan: Stop"
      Timer_Barc_scan_is_counting = False
      $ 340 "If Timer_Barc_scan≥60"
      if (Timer_Barc_scan >= 60):
        $ 341 "set_error(5200)"
        set_error(5200)
      end
    end
  end
  $ 342 "'=========='"
  # '=========='
  $ 343 "PostSettings"
  $ 344 "OBJ_Picked≔rq_is_object_detected()"
  global OBJ_Picked= rq_is_object_detected ()
  $ 345 "If OBJ_Picked"
  if (OBJ_Picked):
    $ 346 "rq_set_force_norm(50)"
     rq_set_force_norm (50)
  end
end
